TYPE ST_BoxConfig :
STRUCT
    sId               : STRING(20);     // slug of the name: lowercase letters, digits and '-'
    sControllerName   : STRING(40);     // exactly the label the website uses for this controller
    nFeedId           : INT := 1;       // index into GVL_Config.aFeeds
    bHasEcPowerSupply : BOOL;           // TRUE: live values come from the EtherCAT supply in the box
    nPixelCount       : UDINT;
    fMaxDcCurrent     : LREAL := 20.0;  // A
    fNominalDcVolts   : LREAL := 24.0;  // turns an estimated share into DC amps
    fPsuEfficiency    : LREAL := 0.95;  // DC power out / AC power in
    fWireLengthFt     : LREAL := 0.0;   // one-way length of the box's AC cable from where it branches off the feed
    nWireAwg          : INT := 12;      // AWG of one conductor, copper
END_STRUCT
END_TYPE

(* stored: Version 1.1.0.1
   DUT ST_BoxConfig: Id {6a2d88ce-d797-411d-902e-cc3ed1de09f3} *)
